TYPE ST_PolarIIChamber_ExhaustServiceParam :
STRUCT
	Fan : ARRAY[1..4] OF ST_PolarIIChamber_ExhaustFanServiceParam;
	Damper : ST_PolarIIChamber_ExhaustDamperServiceParam;
END_STRUCT
END_TYPE

(* stored: Version 1.1.0.1, ProductVersion 3.1.4026.18
   DUT ST_PolarIIChamber_ExhaustServiceParam: Id {14000000-0000-0000-0000-000000000071} *)
